// TIA Portal V21 export
// export: Created 2026-11-10T07:35:24.7972435Z, ExportSetting WithDefaults, DisplayName Totally Integrated Automation Portal, DisplayVersion V21 Update 3, DisplayName STEP 7 Professional, DisplayVersion V21 Update 3, DisplayName STEP 7 Safety, DisplayVersion V21, DisplayName Tech WebApplication, DisplayVersion V21, DisplayName WinCC Basic/Comfort/Advanced, DisplayVersion V21 Update 3, DisplayName WinCC Unified, DisplayVersion V21 Update 3
FUNCTION_BLOCK "FB_Lad_ou001"   // FB194, LAD
{ S7_Optimized_Access := 'TRUE' }
VERSION : 0.1
// stored: AutoNumber true, IsIECCheckEnabled false, IsRetainMemResEnabled false, MemoryReserve 100, SetENOAutomatically false, UDAEnableTagReadback false
   VAR_INPUT
      v_req : Bool;
      v_cont : Bool;
      v_len : UInt;
   END_VAR
   VAR_OUTPUT
      v_done : Bool;
      v_busy : Bool;
      v_error : Bool;
      v_status : Word;
   END_VAR
   VAR_IN_OUT
      v_connect : TCON_Param;
      v_data : Array[0..99] of Byte;
      v_com_rst : Bool;
      v_addr : Variant;
   END_VAR
   VAR
      inst { S7_SetPoint := 'True'} : TSEND_C;
   END_VAR
BEGIN

REGION Network 1: TSEND_C - Send data via Ethernet
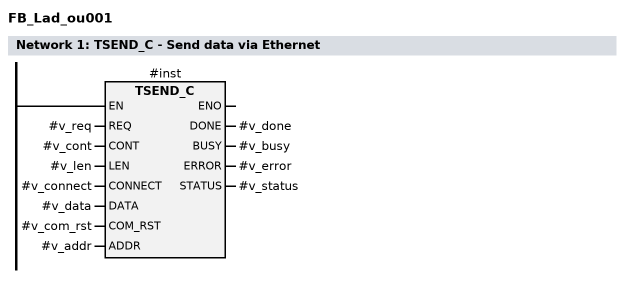
   RUNG wire#powerrail
      #inst.TSEND_C(REQ := #v_req, CONT := #v_cont, LEN := #v_len, CONNECT := #v_connect, DATA := #v_data, COM_RST := #v_com_rst, DONE => #v_done, BUSY => #v_busy, ERROR => #v_error, STATUS => #v_status, ADDR := #v_addr)
   END_RUNG
   // the same network as SCL:
   #inst(REQ := #v_req,   // TSEND_C
         CONT := #v_cont,
         LEN := #v_len,
         CONNECT := #v_connect,
         DATA := #v_data,
         COM_RST := #v_com_rst,
         ADDR := #v_addr,
         DONE => #v_done,
         BUSY => #v_busy,
         ERROR => #v_error,
         STATUS => #v_status);
END_REGION
END_FUNCTION_BLOCK
